Fanuc KAREL source: kb00141.KL

-- PROVISIONAL review KL for V1013-1; original PC SHA256 0dafbf813e8d7be682458d225a008f1f01b90a60276cd4db84a26e96841de0f3
-- Incomplete behavior may be omitted. Consult companion uncertainty JSON. Do not deploy.
PROGRAM KB00141
%NOLOCKGROUP
BEGIN
  -- UNRESOLVED_PC offsets 5-14; opcodes 3F,75
  -- UNRESOLVED_PC offsets 19-26; opcodes 9D,23
  -- UNRESOLVED_PC offsets 31-49; opcodes 27,22,2A,22,31
  -- UNRESOLVED_PC offsets 54-58; opcodes 7F
END KB00141
